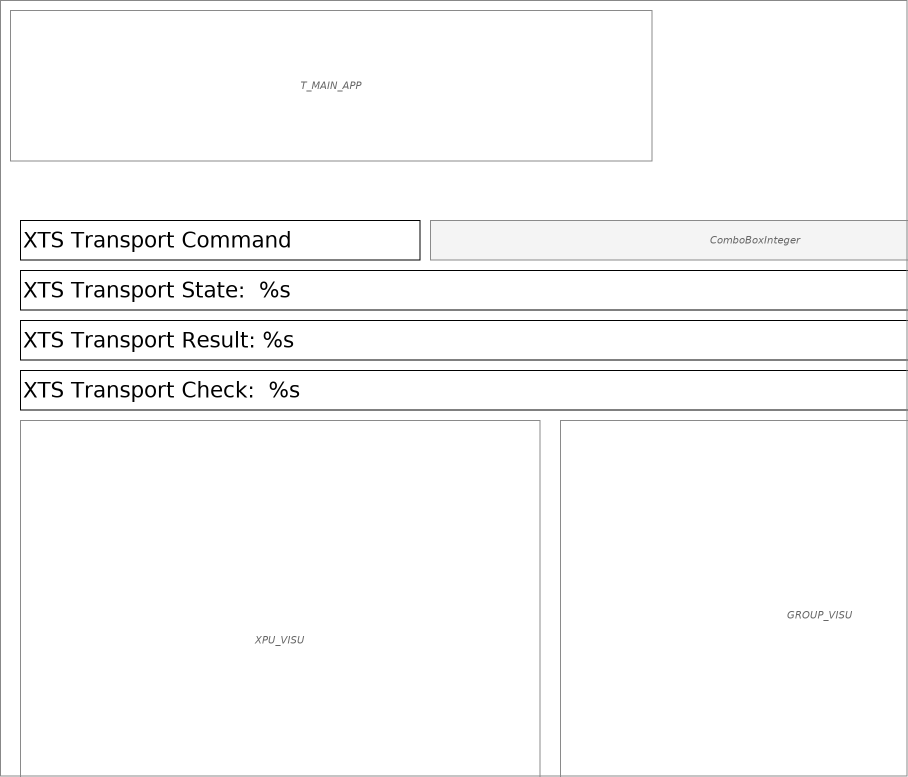
VISUALIZATION VIS_APPLICATION_EXAMPLE  // 908x777
    Group (20,220 888x557)
        Rectangle (0,0 400x40), "XTS Transport Command"
        ComboBoxInteger (410,0 650x40), variable: GVL_XTS.XtsTransportCtrl.Cmd, text list: 'TL_E_CTRL_TRANSPORT'
        Rectangle (0,50 1060x40), "XTS Transport State: %s", text variable: MAIN_XTS.sTransportState
        Rectangle (0,100 1060x40), "XTS Transport Result: %s", text variable: MAIN_XTS.sTransportResult
        Rectangle (0,150 1060x40), "XTS Transport Check: %s", text variable: MAIN_XTS.sTransportCheck
        Frame (0,200 520x440)
            shows XPU_VISU(stXpuState := GVL_XTS.XtsTransportState.XpuState, stXpuInfo := GVL_XTS.XtsTransportState.XpuInfo, stXpuStrings := MAIN_XTS.stXpuStrings)
        Frame (540,200 520x390)
            shows GROUP_VISU(stGroupInfo := GVL_XTS.XtsTransportState.GroupInfo, sGroupState := MAIN_XTS.sCaGroupState)
    Frame (10,10 642x151)
        shows T_MAIN_APP(DataIn := MAIN_APP.stMainVis, DataOut := MAIN_APP.stVisMain)
END_VISUALIZATION

(* stored: Version 1.1.0.1
   Visu VIS_APPLICATION_EXAMPLE: Id {73dd070a-44e9-4cb3-8cdb-da9d7a0d1e0b} *)
